// LS Electric XG5000 project: 555
// PLC LSPLC

PROGRAM E2E_PICKNPLACE (task: 스캔 프로그램)

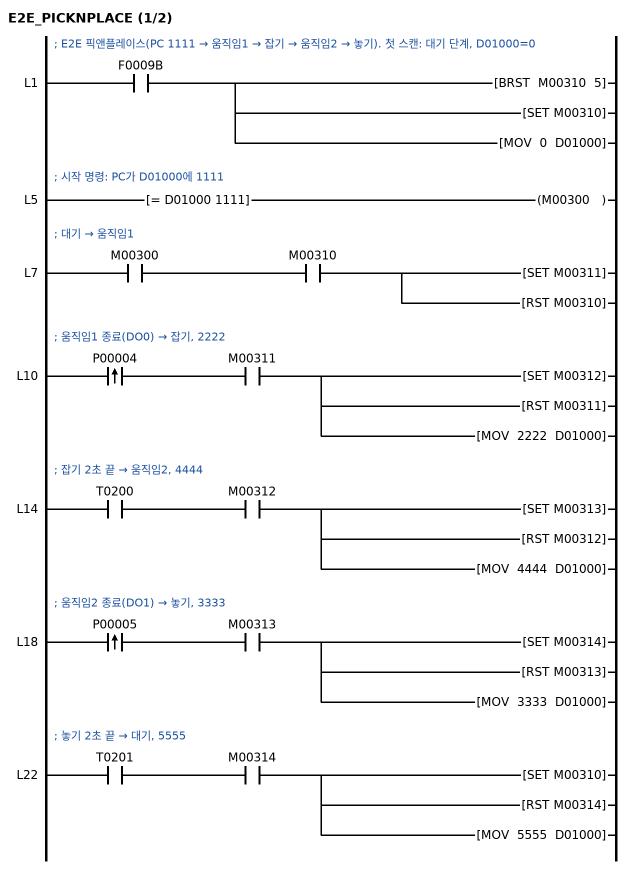
// E2E 픽앤플레이스(PC 1111 → 움직임1 → 잡기 → 움직임2 → 놓기). 첫 스캔: 대기 단계, D01000=0
; L1
LOAD      F0009B
BRST      M00310 5
SET       M00310
MOV       0 D01000
// 시작 명령: PC가 D01000에 1111
; L5
LOAD=     D01000 1111
OUT       M00300
// 대기 → 움직임1
; L7
LOAD      M00300
AND       M00310
SET       M00311
RST       M00310
// 움직임1 종료(DO0) → 잡기, 2222
; L10
LOADP     P00004
AND       M00311
SET       M00312
RST       M00311
MOV       2222 D01000
// 잡기 2초 끝 → 움직임2, 4444
; L14
LOAD      T0200
AND       M00312
SET       M00313
RST       M00312
MOV       4444 D01000
// 움직임2 종료(DO1) → 놓기, 3333
; L18
LOADP     P00005
AND       M00313
SET       M00314
RST       M00313
MOV       3333 D01000
// 놓기 2초 끝 → 대기, 5555
; L22
LOAD      T0201
AND       M00314
SET       M00310
RST       M00314
MOV       5555 D01000

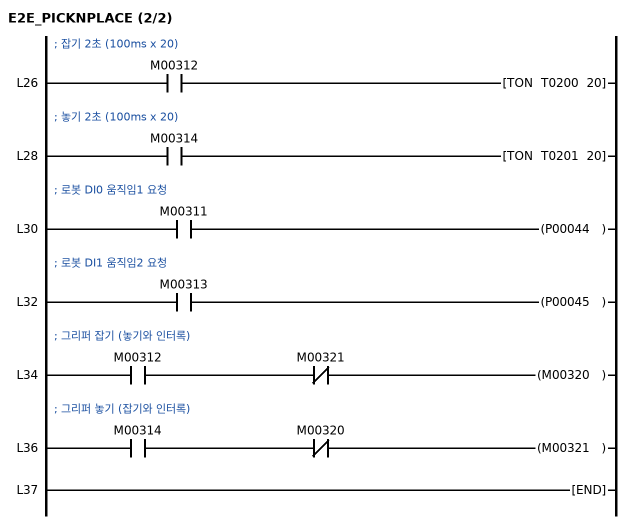
// 잡기 2초 (100ms x 20)
; L26
LOAD      M00312
TON       T0200 20
// 놓기 2초 (100ms x 20)
; L28
LOAD      M00314
TON       T0201 20
// 로봇 DI0 움직임1 요청
; L30
LOAD      M00311
OUT       P00044
// 로봇 DI1 움직임2 요청
; L32
LOAD      M00313
OUT       P00045
// 그리퍼 잡기 (놓기와 인터록)
; L34
LOAD      M00312
AND NOT   M00321
OUT       M00320
// 그리퍼 놓기 (잡기와 인터록)
; L36
LOAD      M00314
AND NOT   M00320
OUT       M00321
; L37
END

VARIABLES AND COMMENTS (devices not used above)
P00041	BIT	GL1
P00000	BIT	PB1
P00001	BIT	PB2
P00042	BIT	YL1
M00103	BIT	상승1
P00007	BIT	상승단
P00046	BIT	승강밸브
M00100	BIT	원점대기
M00102	BIT	잡기대기
T0100	BIT/WORD	타이머_1초
M00101	BIT	하강1
P00008	BIT	하강단